Fanuc KAREL source: kf00114.KL

-- PROVISIONAL review KL for V940-1; original PC SHA256 291bad81a49117034e70037473c7e0eb1799210282e95c76359dbb79d44c14e7
-- Incomplete behavior may be omitted. Consult companion uncertainty JSON. Do not deploy.
PROGRAM KF00114
%NOLOCKGROUP
BEGIN
  -- V9_ZERO_TABLE_METADATA_HINT layout=0001; no indexed target words; source/name/runtime held
  -- V9_CALL_MODE_HINT routine#1 actual=I type=INTEGER mode=address_style
  -- UNRESOLVED_PC offsets 0-1; opcodes 7B
  -- UNRESOLVED_PC offsets 6-20; opcodes 2D,9D,52,23
  -- UNRESOLVED_PC offsets 25-29; opcodes 7F
  -- UNRESOLVED_PC offsets 34-44; opcodes 27,22,AA
  -- UNRESOLVED_PC offsets 49-53; opcodes 7F
END KF00114
